Fanuc KAREL source: KT00682.KL

PROGRAM KT00682
%NOLOCKGROUP
VAR
  P1: JOINTPOS
  P2: JOINTPOS
  OUT: INTEGER
BEGIN
  OUT = + P1
END KT00682
